{region 'Documentation'}
(*!
<summary>Read-only Preparation view; querying does not execute resource actions.</summary>
<description>
This interface exposes only the last reported Status by value. The owner calls the concrete Preparation cyclically with Enable and its resource-specific bindings; the interface provides no generic activation, initialization or reset operation.
</description>
*)
{endregion}
INTERFACE I_Preparation

{region 'Documentation'}
(*!
<summary>Current Preparation status by value; querying does not execute resource actions.</summary>
*)
{endregion}
PROPERTY Status : ST_PreparationStatus //! Current Preparation status by value; querying does not execute resource actions.
GET // PUBLIC
END_GET
END_PROPERTY

END_INTERFACE

(* stored: Version 1.1.0.1
   Itf I_Preparation: Id {d9c504ce-c39f-43a6-9e95-f5b84a6bf3fe}
   Property Status: Id {b8e8978c-7034-47d9-a809-4b4af0330a0f}
   Get Get: Id {128d4400-cd74-4aed-91b6-4380b197bf16} *)
